(* CoDeSys 2.3 export: ld.exp *)

(* POU PLC_LD_PRG_TR, LD *)
PROGRAM PLC_LD_PRG_TR
VAR
END_VAR
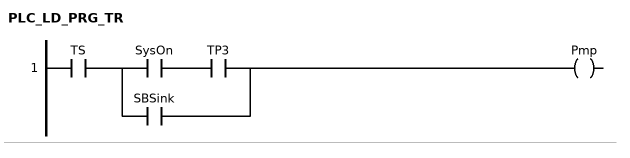
_LD_ (* Ladder Diagram *)
NETWORK 1
	[TS] - { [SysOn] - [TP3] | [SBSink] } --- (Pmp)
_END_LD_
(* the same logic as Structured Text *)
(* Network 1 *)
Pmp := TS AND (SysOn AND TP3 OR SBSink);
END_PROGRAM
